// TIA Portal V20 export
ORGANIZATION_BLOCK "ProgrammingError"   // OB121, LAD, ProgrammingError
TITLE = ProgrammingError
{ S7_Optimized_Access := 'TRUE' }
AUTHOR : IA
FAMILY : PRUEBA
VERSION : 0.1
// Tanda 7: ProgrammingError, incrementa ErroresProg
// stored: IsIECCheckEnabled false, SetENOAutomatically false
   VAR_INPUT
      BlockNr : UInt;
      Reaction : USInt;
      Fault_ID : Byte;
      BlockType : USInt;
      Area : USInt;
      DBNr : DB_ANY;
      Csg_OBNr : OB_ANY;
      Csg_Prio : USInt;
      Width : USInt;
   END_VAR
BEGIN

REGION Network 1: Contador de vida
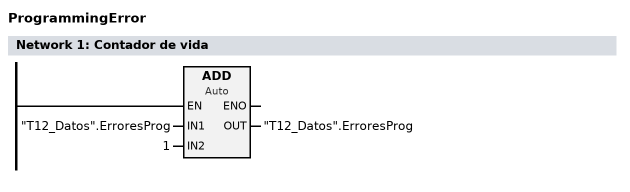
   RUNG wire#powerrail
      Add(in1 := "T12_Datos".ErroresProg, in2 := 1, out => "T12_Datos".ErroresProg)
   END_RUNG
   // the same network as SCL:
   "T12_Datos".ErroresProg := "T12_Datos".ErroresProg + 1;
END_REGION
END_ORGANIZATION_BLOCK
